TYPE ST_PolarIIChamber_ArmServiceParam :
STRUCT
	Lift : ST_PolarIIChamber_LiftTopDownServiceParam;
	Rotate : ST_PolarIIChamber_ArmRotateServiceParam;
	Nozzle : ARRAY[1..3] OF ST_PolarIIChamber_NozzleSupplyServiceParam; // Unsupported array elements are ignored.
	NozzlePort : ST_PolarIIChamber_NozzlePortServiceParam; // Unsupported for Arm3 and Arm4.
END_STRUCT
END_TYPE

(* stored: Version 1.1.0.1, ProductVersion 3.1.4026.18
   DUT ST_PolarIIChamber_ArmServiceParam: Id {14000000-0000-0000-0000-000000000059} *)
